FUNCTION_BLOCK PUMP_STATION (* Migrated from IEC 61131-3 ST *)
  (* Standard: 61499-2 *)
  (* Version 1.0, 2026-11-06, st2fb *)
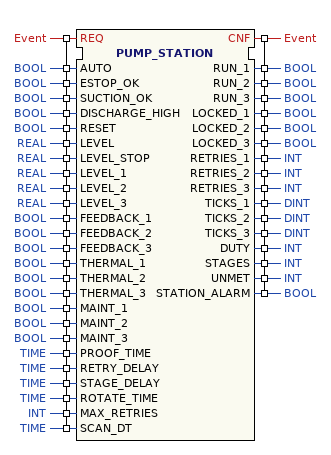
  EVENT_INPUT
    REQ WITH AUTO, ESTOP_OK, SUCTION_OK, DISCHARGE_HIGH, RESET, LEVEL, LEVEL_STOP, LEVEL_1, LEVEL_2, LEVEL_3, FEEDBACK_1, FEEDBACK_2, FEEDBACK_3, THERMAL_1, THERMAL_2, THERMAL_3, MAINT_1, MAINT_2, MAINT_3, PROOF_TIME, RETRY_DELAY, STAGE_DELAY, ROTATE_TIME, MAX_RETRIES, SCAN_DT;
  END_EVENT
  EVENT_OUTPUT
    CNF WITH RUN_1, RUN_2, RUN_3, LOCKED_1, LOCKED_2, LOCKED_3, RETRIES_1, RETRIES_2, RETRIES_3, TICKS_1, TICKS_2, TICKS_3, DUTY, STAGES, UNMET, STATION_ALARM;
  END_EVENT
  VAR_INPUT
    AUTO : BOOL;
    ESTOP_OK : BOOL;
    SUCTION_OK : BOOL;
    DISCHARGE_HIGH : BOOL;
    RESET : BOOL;
    LEVEL : REAL;
    LEVEL_STOP : REAL;
    LEVEL_1 : REAL;
    LEVEL_2 : REAL;
    LEVEL_3 : REAL;
    FEEDBACK_1 : BOOL;
    FEEDBACK_2 : BOOL;
    FEEDBACK_3 : BOOL;
    THERMAL_1 : BOOL;
    THERMAL_2 : BOOL;
    THERMAL_3 : BOOL;
    MAINT_1 : BOOL;
    MAINT_2 : BOOL;
    MAINT_3 : BOOL;
    PROOF_TIME : TIME;
    RETRY_DELAY : TIME;
    STAGE_DELAY : TIME;
    ROTATE_TIME : TIME;
    MAX_RETRIES : INT;
    SCAN_DT : TIME;
  END_VAR
  VAR_OUTPUT
    RUN_1 : BOOL;
    RUN_2 : BOOL;
    RUN_3 : BOOL;
    LOCKED_1 : BOOL;
    LOCKED_2 : BOOL;
    LOCKED_3 : BOOL;
    RETRIES_1 : INT;
    RETRIES_2 : INT;
    RETRIES_3 : INT;
    TICKS_1 : DINT;
    TICKS_2 : DINT;
    TICKS_3 : DINT;
    DUTY : INT;
    STAGES : INT;
    UNMET : INT;
    STATION_ALARM : BOOL;
  END_VAR
  VAR
    ST2FB_NOW : TIME;
    VIEW_AV_1 : BOOL;
    VIEW_AV_2 : BOOL;
    VIEW_AV_3 : BOOL;
    VIEW_TK_1 : DINT;
    VIEW_TK_2 : DINT;
    VIEW_TK_3 : DINT;
    CALLS_1 : BOOL;
    CALLS_2 : BOOL;
    CALLS_3 : BOOL;
    PREF_1 : INT := 1;
    PREF_2 : INT := 2;
    PREF_3 : INT := 3;
    WANTED : INT;
    PERMIT : BOOL;
    ST_IN : BOOL;
    ST_PT : TIME;
    ST_Q : BOOL;
    ST_ET : TIME;
    ST_STATE : INT;
    ST_PREV_IN : BOOL;
    ST_START_TIME : TIME;
    RT_IN : BOOL;
    RT_PT : TIME;
    RT_Q : BOOL;
    RT_ET : TIME;
    RT_STATE : INT;
    RT_PREV_IN : BOOL;
    RT_START_TIME : TIME;
    ALARM_Q1 : BOOL;
    BEST : INT;
    BEST_TICKS : DINT;
    I : INT;
    CANDIDATE : INT;
    REMAIN : INT;
    TMP_AV : BOOL;
    TMP_TK : DINT;
    TMP_IDX : INT;
    U1_STATE : INT;
    U1_FAILED : BOOL;
    U1_RUN : BOOL;
    U1_AVAILABLE : BOOL;
    U1_LOCKED : BOOL;
    U1_RETRIES : INT;
    U1_TICKS : DINT;
    U1_PR_IN : BOOL;
    U1_PR_PT : TIME;
    U1_PR_Q : BOOL;
    U1_PR_ET : TIME;
    U1_PR_STATE : INT;
    U1_PR_PREV_IN : BOOL;
    U1_PR_START_TIME : TIME;
    U1_HO_IN : BOOL;
    U1_HO_PT : TIME;
    U1_HO_Q : BOOL;
    U1_HO_ET : TIME;
    U1_HO_STATE : INT;
    U1_HO_PREV_IN : BOOL;
    U1_HO_START_TIME : TIME;
    U2_STATE : INT;
    U2_FAILED : BOOL;
    U2_RUN : BOOL;
    U2_AVAILABLE : BOOL;
    U2_LOCKED : BOOL;
    U2_RETRIES : INT;
    U2_TICKS : DINT;
    U2_PR_IN : BOOL;
    U2_PR_PT : TIME;
    U2_PR_Q : BOOL;
    U2_PR_ET : TIME;
    U2_PR_STATE : INT;
    U2_PR_PREV_IN : BOOL;
    U2_PR_START_TIME : TIME;
    U2_HO_IN : BOOL;
    U2_HO_PT : TIME;
    U2_HO_Q : BOOL;
    U2_HO_ET : TIME;
    U2_HO_STATE : INT;
    U2_HO_PREV_IN : BOOL;
    U2_HO_START_TIME : TIME;
    U3_STATE : INT;
    U3_FAILED : BOOL;
    U3_RUN : BOOL;
    U3_AVAILABLE : BOOL;
    U3_LOCKED : BOOL;
    U3_RETRIES : INT;
    U3_TICKS : DINT;
    U3_PR_IN : BOOL;
    U3_PR_PT : TIME;
    U3_PR_Q : BOOL;
    U3_PR_ET : TIME;
    U3_PR_STATE : INT;
    U3_PR_PREV_IN : BOOL;
    U3_PR_START_TIME : TIME;
    U3_HO_IN : BOOL;
    U3_HO_PT : TIME;
    U3_HO_Q : BOOL;
    U3_HO_ET : TIME;
    U3_HO_STATE : INT;
    U3_HO_PREV_IN : BOOL;
    U3_HO_START_TIME : TIME;
  END_VAR
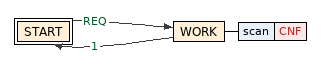
  EC_STATES
    START;
    WORK : scan -> CNF;
  END_STATES
  EC_TRANSITIONS
    START TO WORK := REQ;
    WORK TO START := 1;
  END_TRANSITIONS
  ALGORITHM scan IN ST:
ST2FB_NOW := ST2FB_NOW + SCAN_DT;
PERMIT := ESTOP_OK AND SUCTION_OK AND NOT DISCHARGE_HIGH;

IF NOT AUTO OR LEVEL <= LEVEL_STOP THEN
  WANTED := 0;
ELSIF LEVEL >= LEVEL_3 THEN
  WANTED := 3;
ELSIF LEVEL >= LEVEL_2 THEN
  WANTED := MAX(WANTED, 2);
ELSIF LEVEL >= LEVEL_1 THEN
  WANTED := MAX(WANTED, 1);
END_IF;

ST_IN := (STAGES < WANTED) AND NOT ST_Q;
ST_PT := STAGE_DELAY;
IF (ST_STATE = 0) AND NOT ST_PREV_IN AND ST_IN THEN
  ST_STATE := 1;
  ST_Q := FALSE;
  ST_START_TIME := ST2FB_NOW;
ELSE
  IF NOT ST_IN THEN
    ST_ET := T#0s;
    ST_Q := FALSE;
    ST_STATE := 0;
  ELSIF ST_STATE = 1 THEN
    IF ST_START_TIME + ST_PT <= ST2FB_NOW THEN
      ST_STATE := 2;
      ST_Q := TRUE;
      ST_ET := ST_PT;
    ELSE
      ST_ET := ST2FB_NOW - ST_START_TIME;
    END_IF;
  END_IF;
END_IF;
ST_PREV_IN := ST_IN;

IF STAGES > WANTED THEN
  STAGES := WANTED;
ELSIF ST_Q THEN
  STAGES := STAGES + 1;
END_IF;

RT_IN := AUTO AND NOT RT_Q;
RT_PT := ROTATE_TIME;
IF (RT_STATE = 0) AND NOT RT_PREV_IN AND RT_IN THEN
  RT_STATE := 1;
  RT_Q := FALSE;
  RT_START_TIME := ST2FB_NOW;
ELSE
  IF NOT RT_IN THEN
    RT_ET := T#0s;
    RT_Q := FALSE;
    RT_STATE := 0;
  ELSIF RT_STATE = 1 THEN
    IF RT_START_TIME + RT_PT <= ST2FB_NOW THEN
      RT_STATE := 2;
      RT_Q := TRUE;
      RT_ET := RT_PT;
    ELSE
      RT_ET := ST2FB_NOW - RT_START_TIME;
    END_IF;
  END_IF;
END_IF;
RT_PREV_IN := RT_IN;

TMP_IDX := MAX(DUTY, 1);
IF TMP_IDX = 1 THEN
  TMP_AV := VIEW_AV_1;
ELSIF TMP_IDX = 2 THEN
  TMP_AV := VIEW_AV_2;
ELSE
  TMP_AV := VIEW_AV_3;
END_IF;
IF RT_Q OR (DUTY = 0) OR NOT TMP_AV THEN
  BEST := 0;
  BEST_TICKS := 2147483647;
  FOR I := 1 TO 3 DO
    IF I = 1 THEN
      CANDIDATE := PREF_1;
    ELSIF I = 2 THEN
      CANDIDATE := PREF_2;
    ELSE
      CANDIDATE := PREF_3;
    END_IF;
    IF CANDIDATE = 1 THEN
      TMP_AV := VIEW_AV_1;
      TMP_TK := VIEW_TK_1;
    ELSIF CANDIDATE = 2 THEN
      TMP_AV := VIEW_AV_2;
      TMP_TK := VIEW_TK_2;
    ELSE
      TMP_AV := VIEW_AV_3;
      TMP_TK := VIEW_TK_3;
    END_IF;
    IF TMP_AV AND (TMP_TK < BEST_TICKS) THEN
      BEST := CANDIDATE;
      BEST_TICKS := TMP_TK;
    END_IF;
  END_FOR;
  IF BEST <> 0 THEN
    DUTY := BEST;
  END_IF;
END_IF;

CALLS_1 := FALSE;
CALLS_2 := FALSE;
CALLS_3 := FALSE;
REMAIN := STAGES;
FOR I := 0 TO 2 DO
  IF REMAIN <> 0 THEN
    CANDIDATE := (MAX(DUTY, 1) + I - 1) MOD 3 + 1;
    IF CANDIDATE = 1 THEN
      TMP_AV := VIEW_AV_1;
    ELSIF CANDIDATE = 2 THEN
      TMP_AV := VIEW_AV_2;
    ELSE
      TMP_AV := VIEW_AV_3;
    END_IF;
    IF TMP_AV THEN
      IF CANDIDATE = 1 THEN
        CALLS_1 := TRUE;
      ELSIF CANDIDATE = 2 THEN
        CALLS_2 := TRUE;
      ELSE
        CALLS_3 := TRUE;
      END_IF;
      REMAIN := REMAIN - 1;
    END_IF;
  END_IF;
END_FOR;
UNMET := REMAIN;

(* pump 1 *)
IF RESET AND NOT THERMAL_1 THEN
  U1_RETRIES := 0;
  IF U1_STATE = 4 THEN
    U1_STATE := 0;
  END_IF;
END_IF;
IF NOT PERMIT AND U1_STATE <> 4 THEN
  U1_STATE := 0;
END_IF;
U1_FAILED := FALSE;
CASE U1_STATE OF
  0:
    IF CALLS_1 AND PERMIT AND NOT MAINT_1 AND NOT THERMAL_1 THEN
      U1_STATE := 1;
    END_IF;
  1:
    IF NOT CALLS_1 THEN
      U1_STATE := 0;
    ELSIF THERMAL_1 OR U1_PR_Q THEN
      U1_FAILED := TRUE;
    ELSIF FEEDBACK_1 THEN
      U1_STATE := 2;
    END_IF;
  2:
    IF NOT CALLS_1 THEN
      U1_STATE := 0;
    ELSIF THERMAL_1 OR NOT FEEDBACK_1 THEN
      U1_FAILED := TRUE;
    END_IF;
  3:
    IF U1_HO_Q THEN
      U1_STATE := 0;
    END_IF;
END_CASE;
IF U1_FAILED THEN
  U1_RETRIES := U1_RETRIES + 1;
  IF U1_RETRIES >= MAX_RETRIES THEN
    U1_STATE := 4;
  ELSE
    U1_STATE := 3;
  END_IF;
END_IF;
U1_PR_IN := U1_STATE = 1;
U1_PR_PT := PROOF_TIME;
IF (U1_PR_STATE = 0) AND NOT U1_PR_PREV_IN AND U1_PR_IN THEN
  U1_PR_STATE := 1;
  U1_PR_Q := FALSE;
  U1_PR_START_TIME := ST2FB_NOW;
ELSE
  IF NOT U1_PR_IN THEN
    U1_PR_ET := T#0s;
    U1_PR_Q := FALSE;
    U1_PR_STATE := 0;
  ELSIF U1_PR_STATE = 1 THEN
    IF U1_PR_START_TIME + U1_PR_PT <= ST2FB_NOW THEN
      U1_PR_STATE := 2;
      U1_PR_Q := TRUE;
      U1_PR_ET := U1_PR_PT;
    ELSE
      U1_PR_ET := ST2FB_NOW - U1_PR_START_TIME;
    END_IF;
  END_IF;
END_IF;
U1_PR_PREV_IN := U1_PR_IN;
U1_HO_IN := U1_STATE = 3;
U1_HO_PT := RETRY_DELAY;
IF (U1_HO_STATE = 0) AND NOT U1_HO_PREV_IN AND U1_HO_IN THEN
  U1_HO_STATE := 1;
  U1_HO_Q := FALSE;
  U1_HO_START_TIME := ST2FB_NOW;
ELSE
  IF NOT U1_HO_IN THEN
    U1_HO_ET := T#0s;
    U1_HO_Q := FALSE;
    U1_HO_STATE := 0;
  ELSIF U1_HO_STATE = 1 THEN
    IF U1_HO_START_TIME + U1_HO_PT <= ST2FB_NOW THEN
      U1_HO_STATE := 2;
      U1_HO_Q := TRUE;
      U1_HO_ET := U1_HO_PT;
    ELSE
      U1_HO_ET := ST2FB_NOW - U1_HO_START_TIME;
    END_IF;
  END_IF;
END_IF;
U1_HO_PREV_IN := U1_HO_IN;
U1_RUN := (U1_STATE = 1) OR (U1_STATE = 2);
U1_AVAILABLE := NOT MAINT_1 AND NOT THERMAL_1 AND (U1_STATE <> 3) AND (U1_STATE <> 4);
U1_LOCKED := U1_STATE = 4;
IF U1_STATE = 2 THEN
  U1_TICKS := U1_TICKS + 1;
END_IF;

(* pump 2 *)
IF RESET AND NOT THERMAL_2 THEN
  U2_RETRIES := 0;
  IF U2_STATE = 4 THEN
    U2_STATE := 0;
  END_IF;
END_IF;
IF NOT PERMIT AND U2_STATE <> 4 THEN
  U2_STATE := 0;
END_IF;
U2_FAILED := FALSE;
CASE U2_STATE OF
  0:
    IF CALLS_2 AND PERMIT AND NOT MAINT_2 AND NOT THERMAL_2 THEN
      U2_STATE := 1;
    END_IF;
  1:
    IF NOT CALLS_2 THEN
      U2_STATE := 0;
    ELSIF THERMAL_2 OR U2_PR_Q THEN
      U2_FAILED := TRUE;
    ELSIF FEEDBACK_2 THEN
      U2_STATE := 2;
    END_IF;
  2:
    IF NOT CALLS_2 THEN
      U2_STATE := 0;
    ELSIF THERMAL_2 OR NOT FEEDBACK_2 THEN
      U2_FAILED := TRUE;
    END_IF;
  3:
    IF U2_HO_Q THEN
      U2_STATE := 0;
    END_IF;
END_CASE;
IF U2_FAILED THEN
  U2_RETRIES := U2_RETRIES + 1;
  IF U2_RETRIES >= MAX_RETRIES THEN
    U2_STATE := 4;
  ELSE
    U2_STATE := 3;
  END_IF;
END_IF;
U2_PR_IN := U2_STATE = 1;
U2_PR_PT := PROOF_TIME;
IF (U2_PR_STATE = 0) AND NOT U2_PR_PREV_IN AND U2_PR_IN THEN
  U2_PR_STATE := 1;
  U2_PR_Q := FALSE;
  U2_PR_START_TIME := ST2FB_NOW;
ELSE
  IF NOT U2_PR_IN THEN
    U2_PR_ET := T#0s;
    U2_PR_Q := FALSE;
    U2_PR_STATE := 0;
  ELSIF U2_PR_STATE = 1 THEN
    IF U2_PR_START_TIME + U2_PR_PT <= ST2FB_NOW THEN
      U2_PR_STATE := 2;
      U2_PR_Q := TRUE;
      U2_PR_ET := U2_PR_PT;
    ELSE
      U2_PR_ET := ST2FB_NOW - U2_PR_START_TIME;
    END_IF;
  END_IF;
END_IF;
U2_PR_PREV_IN := U2_PR_IN;
U2_HO_IN := U2_STATE = 3;
U2_HO_PT := RETRY_DELAY;
IF (U2_HO_STATE = 0) AND NOT U2_HO_PREV_IN AND U2_HO_IN THEN
  U2_HO_STATE := 1;
  U2_HO_Q := FALSE;
  U2_HO_START_TIME := ST2FB_NOW;
ELSE
  IF NOT U2_HO_IN THEN
    U2_HO_ET := T#0s;
    U2_HO_Q := FALSE;
    U2_HO_STATE := 0;
  ELSIF U2_HO_STATE = 1 THEN
    IF U2_HO_START_TIME + U2_HO_PT <= ST2FB_NOW THEN
      U2_HO_STATE := 2;
      U2_HO_Q := TRUE;
      U2_HO_ET := U2_HO_PT;
    ELSE
      U2_HO_ET := ST2FB_NOW - U2_HO_START_TIME;
    END_IF;
  END_IF;
END_IF;
U2_HO_PREV_IN := U2_HO_IN;
U2_RUN := (U2_STATE = 1) OR (U2_STATE = 2);
U2_AVAILABLE := NOT MAINT_2 AND NOT THERMAL_2 AND (U2_STATE <> 3) AND (U2_STATE <> 4);
U2_LOCKED := U2_STATE = 4;
IF U2_STATE = 2 THEN
  U2_TICKS := U2_TICKS + 1;
END_IF;

(* pump 3 *)
IF RESET AND NOT THERMAL_3 THEN
  U3_RETRIES := 0;
  IF U3_STATE = 4 THEN
    U3_STATE := 0;
  END_IF;
END_IF;
IF NOT PERMIT AND U3_STATE <> 4 THEN
  U3_STATE := 0;
END_IF;
U3_FAILED := FALSE;
CASE U3_STATE OF
  0:
    IF CALLS_3 AND PERMIT AND NOT MAINT_3 AND NOT THERMAL_3 THEN
      U3_STATE := 1;
    END_IF;
  1:
    IF NOT CALLS_3 THEN
      U3_STATE := 0;
    ELSIF THERMAL_3 OR U3_PR_Q THEN
      U3_FAILED := TRUE;
    ELSIF FEEDBACK_3 THEN
      U3_STATE := 2;
    END_IF;
  2:
    IF NOT CALLS_3 THEN
      U3_STATE := 0;
    ELSIF THERMAL_3 OR NOT FEEDBACK_3 THEN
      U3_FAILED := TRUE;
    END_IF;
  3:
    IF U3_HO_Q THEN
      U3_STATE := 0;
    END_IF;
END_CASE;
IF U3_FAILED THEN
  U3_RETRIES := U3_RETRIES + 1;
  IF U3_RETRIES >= MAX_RETRIES THEN
    U3_STATE := 4;
  ELSE
    U3_STATE := 3;
  END_IF;
END_IF;
U3_PR_IN := U3_STATE = 1;
U3_PR_PT := PROOF_TIME;
IF (U3_PR_STATE = 0) AND NOT U3_PR_PREV_IN AND U3_PR_IN THEN
  U3_PR_STATE := 1;
  U3_PR_Q := FALSE;
  U3_PR_START_TIME := ST2FB_NOW;
ELSE
  IF NOT U3_PR_IN THEN
    U3_PR_ET := T#0s;
    U3_PR_Q := FALSE;
    U3_PR_STATE := 0;
  ELSIF U3_PR_STATE = 1 THEN
    IF U3_PR_START_TIME + U3_PR_PT <= ST2FB_NOW THEN
      U3_PR_STATE := 2;
      U3_PR_Q := TRUE;
      U3_PR_ET := U3_PR_PT;
    ELSE
      U3_PR_ET := ST2FB_NOW - U3_PR_START_TIME;
    END_IF;
  END_IF;
END_IF;
U3_PR_PREV_IN := U3_PR_IN;
U3_HO_IN := U3_STATE = 3;
U3_HO_PT := RETRY_DELAY;
IF (U3_HO_STATE = 0) AND NOT U3_HO_PREV_IN AND U3_HO_IN THEN
  U3_HO_STATE := 1;
  U3_HO_Q := FALSE;
  U3_HO_START_TIME := ST2FB_NOW;
ELSE
  IF NOT U3_HO_IN THEN
    U3_HO_ET := T#0s;
    U3_HO_Q := FALSE;
    U3_HO_STATE := 0;
  ELSIF U3_HO_STATE = 1 THEN
    IF U3_HO_START_TIME + U3_HO_PT <= ST2FB_NOW THEN
      U3_HO_STATE := 2;
      U3_HO_Q := TRUE;
      U3_HO_ET := U3_HO_PT;
    ELSE
      U3_HO_ET := ST2FB_NOW - U3_HO_START_TIME;
    END_IF;
  END_IF;
END_IF;
U3_HO_PREV_IN := U3_HO_IN;
U3_RUN := (U3_STATE = 1) OR (U3_STATE = 2);
U3_AVAILABLE := NOT MAINT_3 AND NOT THERMAL_3 AND (U3_STATE <> 3) AND (U3_STATE <> 4);
U3_LOCKED := U3_STATE = 4;
IF U3_STATE = 2 THEN
  U3_TICKS := U3_TICKS + 1;
END_IF;

VIEW_AV_1 := U1_AVAILABLE;
VIEW_TK_1 := U1_TICKS;
VIEW_AV_2 := U2_AVAILABLE;
VIEW_TK_2 := U2_TICKS;
VIEW_AV_3 := U3_AVAILABLE;
VIEW_TK_3 := U3_TICKS;

RUN_1 := U1_RUN;
RUN_2 := U2_RUN;
RUN_3 := U3_RUN;
LOCKED_1 := U1_LOCKED;
LOCKED_2 := U2_LOCKED;
LOCKED_3 := U3_LOCKED;
RETRIES_1 := U1_RETRIES;
RETRIES_2 := U2_RETRIES;
RETRIES_3 := U3_RETRIES;
TICKS_1 := U1_TICKS;
TICKS_2 := U2_TICKS;
TICKS_3 := U3_TICKS;

ALARM_Q1 := (U1_LOCKED OR U2_LOCKED OR U3_LOCKED OR ((UNMET > 0) AND PERMIT)) OR (NOT RESET AND ALARM_Q1);
STATION_ALARM := ALARM_Q1;
  END_ALGORITHM
END_FUNCTION_BLOCK
